(* IEC 61131-3 sources: codesys-api/examples/mqtt_large_payload/st/edge, 3 files *)

(* ---- FB_EdgeReceiver.st ---- *)
FUNCTION_BLOCK FB_EdgeReceiver IMPLEMENTS MQTT.MQTT_SUBSCRIBE_CALLBACK
// Subscription callback for EdgeTest: the size and Adler-32 of the last message, and how many arrived.
// ReceivedCount changes last, so a reader that sees a new count also sees that message's size and sum.
VAR_OUTPUT
	ReceivedCount : UDINT;
	LastSize : UDINT;
	LastAdler32 : UDINT;
	// Messages starting with 8 ASCII digits carry a sequence number (qos_test.py); write ResetSequence online
	LastSequence : UDINT;
	InOrderCount : UDINT;               // sequence = previous + 1
	DuplicateCount : UDINT;             // sequence <= previous: delivered again
	GapCount : UDINT;                   // sequence numbers skipped: lost
END_VAR
VAR_INPUT
	ResetSequence : BOOL;               // written online; cleared by the next message
END_VAR
// ---- implementation ----

(* ---- EdgeTest.st ---- *)
PROGRAM EdgeTest
// Edge-case test for the MQTT library, driven online by edge_test.py; idle unless IsEnabled.
// Send: when SendSequence changes, publishes SendSize payload bytes on TopicOut. Byte i is
// (i * 31 + SendSequence) MOD 251, so the broker-side checker can verify every byte of every size.
// Receive: every message on TopicIn is counted with its size and Adler-32 (Receiver).
VAR
	IsEnabled : BOOL;                   // written online
	SendSize : UDINT := 100;            // written online: payload bytes of the next message
	IsQos1 : BOOL;                      // written online
	IsQos2 : BOOL;                      // written online: publish at QoS 2 (wins over IsQos1)
	SubscribeQoS : BYTE := 1;           // written online: 0, 1 or 2; takes effect at the next subscribe
	                                    // (qos_test.py switches IsEnabled off and on to resubscribe)
	SendSequence : UDINT;               // written online; a new value starts a send
	DoneSequence : UDINT;               // the sequence of the last message the library reported done
	TimeoutCount : UDINT;               // rising edges of Publisher.SendTimeout
	RejectedCount : UDINT;              // messages the library gave up because the broker refused them
	IsEchoEnabled : BOOL;               // written online: answer every received message on TopicEcho (QoS 1)
	EchoCount : UDINT;                  // echoes the library reported done
	Receiver : FB_EdgeReceiver;
	TopicEcho : STRING(64) := 'raw_data_demo/edge_echo';
	EchoText : STRING(32);
	EchoPublisher : MQTT.MQTTPublish;
	IsEchoRequested : BOOL;
	IsEchoArmed : BOOL := TRUE;
	EchoedCount : UDINT;                // Receiver.ReceivedCount at the last echo started
	TopicOut : STRING(64) := 'raw_data_demo/edge';
	TopicIn : STRING(64) := 'raw_data_demo/edge_in';
	Publisher : MQTT.MQTTPublish;
	Subscriber : MQTT.MQTTSubscribe;
	IsReady : BOOL;
	IsRequested : BOOL;
	IsArmed : BOOL := TRUE;
	StartedSequence : UDINT;
	RequestSize : UDINT;                // SendSize when the current request started
	PublishQoS : MQTT.QoS;
	SubscribeQoSValue : MQTT.QoS;
	TimeoutEdge : R_TRIG;
	Payload : ARRAY[0..MAX_PAYLOAD - 1] OF BYTE;
	Index : UDINT;
END_VAR
VAR CONSTANT
	MAX_PAYLOAD : UDINT := 40000;
END_VAR
// ---- implementation ----
IF NOT IsReady THEN
	IsReady := TRUE;
	Publisher.SetMqttInOut(MQTT_IN_OUT := PLC_PRG.MqttLink);
	Subscriber.SetMqttInOut(MQTT_IN_OUT := PLC_PRG.MqttLink);
	EchoPublisher.SetMqttInOut(MQTT_IN_OUT := PLC_PRG.MqttLink);
END_IF

CASE SubscribeQoS OF
	0: SubscribeQoSValue := MQTT.QoS.AtMostOnce;
	2: SubscribeQoSValue := MQTT.QoS.ExactlyOnce;
ELSE
	SubscribeQoSValue := MQTT.QoS.AtLeastOnce;
END_CASE
Subscriber(Subscribe := IsEnabled, Topic := ADR(TopicIn), QoSSubscribe := SubscribeQoSValue,
	ExpectingString := FALSE, Callback := Receiver);

// MQTTPublish starts on a rising edge of send: a new request only once the publisher has been called with
// send FALSE after the previous done (IsArmed). Without it a request written in the scan after done is lost.
IF IsEnabled AND NOT IsRequested AND IsArmed AND SendSequence <> StartedSequence AND SendSize > 0 AND SendSize <= MAX_PAYLOAD THEN
	RequestSize := SendSize;	// latched: the publish uses the size this request started with
	FOR Index := 0 TO RequestSize - 1 DO
		Payload[Index] := UDINT_TO_BYTE((Index * 31 + SendSequence) MOD 251);
	END_FOR
	StartedSequence := SendSequence;
	IsRequested := TRUE;
	IsArmed := FALSE;
END_IF
IF IsQos2 THEN
	PublishQoS := MQTT.QoS.ExactlyOnce;
ELSIF IsQos1 THEN
	PublishQoS := MQTT.QoS.AtLeastOnce;
ELSE
	PublishQoS := MQTT.QoS.AtMostOnce;
END_IF
Publisher(Topic := ADR(TopicOut), PublishAsString := FALSE, Payload := ADR(Payload), PayloadLength := RequestSize,
	QoSIn := PublishQoS, MRetain := FALSE, send := IsRequested);
IF NOT IsRequested THEN
	IsArmed := TRUE;	// the publisher has seen send FALSE
END_IF
IF Publisher.done THEN
	IsRequested := FALSE;
	DoneSequence := StartedSequence;
END_IF
// the broker refused the message (it closed the connection after it, three times): given up, not done
IF Publisher.Rejected AND IsRequested THEN
	IsRequested := FALSE;
	RejectedCount := RejectedCount + 1;
END_IF
TimeoutEdge(CLK := Publisher.SendTimeout);
IF TimeoutEdge.Q THEN
	TimeoutCount := TimeoutCount + 1;
END_IF

// Echo (command and acknowledgement round trip): answer the newest received message with its count, QoS 1,
// like PRG_Comms acknowledging a command. Same armed rule as above.
IF IsEchoEnabled AND NOT IsEchoRequested AND IsEchoArmed AND Receiver.ReceivedCount <> EchoedCount THEN
	EchoedCount := Receiver.ReceivedCount;
	EchoText := UDINT_TO_STRING(EchoedCount);
	IsEchoRequested := TRUE;
	IsEchoArmed := FALSE;
END_IF
EchoPublisher(Topic := ADR(TopicEcho), PayloadString := ADR(EchoText), PublishAsString := TRUE,
	QoSIn := MQTT.QoS.AtLeastOnce, MRetain := FALSE, send := IsEchoRequested);
IF NOT IsEchoRequested THEN
	IsEchoArmed := TRUE;
END_IF
IF EchoPublisher.done THEN
	IsEchoRequested := FALSE;
	EchoCount := EchoCount + 1;
END_IF

(* ---- FB_EdgeReceiver.PublishReceived.st ---- *)
METHOD PublishReceived : BOOL
VAR_INPUT
	Data : MQTT.CALLBACK_DATA;
END_VAR
VAR
	Index : UDINT;
	SumA : UDINT;
	SumB : UDINT;
	pByte : POINTER TO BYTE;
	Sequence : UDINT;
	IsSequenced : BOOL;
END_VAR
// ---- implementation ----
// Adler-32 (as zlib.adler32) over the binary payload; the library reuses its buffer after this call.
SumA := 1;
SumB := 0;
pByte := Data.Payload;
IF Data.PayloadSize > 0 AND pByte <> 0 THEN
	FOR Index := 0 TO Data.PayloadSize - 1 DO
		SumA := (SumA + pByte[Index]) MOD 65521;
		SumB := (SumB + SumA) MOD 65521;
	END_FOR
END_IF
LastSize := Data.PayloadSize;
LastAdler32 := SumB * 65536 + SumA;

// Sequence check: 8 leading ASCII digits
IsSequenced := Data.PayloadSize >= 8 AND pByte <> 0;
Sequence := 0;
IF IsSequenced THEN
	FOR Index := 0 TO 7 DO
		IF pByte[Index] < 48 OR pByte[Index] > 57 THEN
			IsSequenced := FALSE;
		ELSE
			Sequence := Sequence * 10 + (pByte[Index] - 48);
		END_IF
	END_FOR
END_IF
IF IsSequenced THEN
	IF ResetSequence THEN
		ResetSequence := FALSE;
		LastSequence := 0;
		InOrderCount := 0;
		DuplicateCount := 0;
		GapCount := 0;
	END_IF
	IF Sequence = LastSequence + 1 THEN
		InOrderCount := InOrderCount + 1;
	ELSIF Sequence <= LastSequence THEN
		DuplicateCount := DuplicateCount + 1;
	ELSE
		GapCount := GapCount + (Sequence - LastSequence - 1);
		InOrderCount := InOrderCount + 1;
	END_IF
	IF Sequence > LastSequence THEN
		LastSequence := Sequence;
	END_IF
END_IF
ReceivedCount := ReceivedCount + 1;
PublishReceived := TRUE;
